Fanuc KAREL source: KA00127.KL

PROGRAM KA00127
%NOLOCKGROUP
VAR
  SRC: ARRAY[2] OF BYTE
  DST: XYZWPREXT
BEGIN
  SRC[1] = 2
  DST = SRC[1]
END KA00127
